(* IEC 61131-3 sources: avi-aoi-management/scripts/ai-eval/ngau-nhien/kho/st-tt3-tre-tru/khung/src, 1 file *)

(* ---- TreTru.st ---- *)
FUNCTION_BLOCK TreTru
VAR_INPUT
    PV : REAL;
    SP : REAL;
    DAI : REAL;
    CHE_DO_LAM_LANH : BOOL;
END_VAR
VAR_OUTPUT
    Q : BOOL;
END_VAR
    (* TODO: cài đặt theo đề bài *)
    Q := FALSE;
END_FUNCTION_BLOCK
